SUBAPPLICATION INI_IN_AND_STORE_AUI2 (* INI Laden und Speichern von AUI2-Daten (reine Ganzzahl 0-N, kein Scale/Decimals) mit zusaetzlichem VALUEO (AUI, plain) fuer einen weiteren Consumer - analog INI_IN_AND_STORE_AUDI2, aber ueber den bidirektionalen AUI2-Adapter (UINT) statt AUDI2 (UDINT), z.B. fuer K eines AOption_AUI_DEMUX_N. *)
  (* Standard: 61499-2; Description: Copyright (c) 2026 Meisterschulen am Ostbahnhof This program and the accompanying materials are made available under the terms of the Eclipse Public License 2.0 which is available at https://www.eclipse.org/legal/epl-2.0/ SPDX-License-Identifier: EPL-2.0 *)
  (* Version 1.0, 2026-10-13, Franz Höpfinger, Meisterschulen am Ostbahnhof, UINT/AUI2-Pendant zu MyLib::sys::INI_IN_AND_STORE_AUDI2: NumericValue_IDA + AD_TO_AUI + AUI_TO_AUI2 + INI_AUI2 (bidirektionaler Adapter statt AUI+Split-Paar), AUI_TO_AUI2.AUI_OUT gesplittet auf Q_NumericValue_AUDI (VT-Anzeige, via AUI_TO_AUDI) und VALUEO (weiterer Consumer, z.B. AOption_AUI_DEMUX_N.K). Strukturell identisch zu INI_IN_AND_STORE_AUDI2, nur mit AUI2 statt AUDI2. *)
  PACKAGE MyLib::sys;
  IMPORT isobus::UT::Q::const::IDs::ID_NULL;
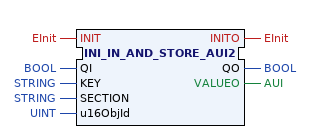
  EVENT_INPUT
    INIT : EInit; (* Initialization Request *)
  END_EVENT
  EVENT_OUTPUT
    INITO : EInit; (* Initialization Confirm *)
  END_EVENT
  VAR_INPUT
    QI : BOOL := TRUE; (* Quality Input - TRUE to enable service *)
    KEY : STRING; (* Key name. *)
    SECTION : STRING; (* Section name. *)
    u16ObjId : UINT := ID_NULL;
  END_VAR
  VAR_OUTPUT
    QO : BOOL; (* Quality Output - TRUE if service executed successfully *)
  END_VAR
  PLUGS
    VALUEO : adapter::types::unidirectional::AUI;
  END_PLUGS
  (* SETM=TRUE - der Boot-Wert laedt so oder so automatisch (INIT -> INITO -> GET -> GETO, unabhaengig von SETM). SETM=TRUE sorgt dafuer, dass auch eine LIVE-Aenderung waehrend des laufenden Betriebs sofort bestaetigt/zurueckgemeldet wird - wichtig, falls der frische Wert noch im selben Lauf weiterverwendet werden soll (z.B. hier ueber VALUEO). *)
  FBS
    ID : isobus::UT::io::NumericValue::NumericValue_IDA;
    AD_TO_AUI : adapter::conversion::unidirectional::AD_TO_AUI;
    AUI_TO_AUI2 : adapter::conversion::bidirectional::AUI_TO_AUI2;
    INI_AUI2 : eclipse4diac::storage::INI_AUI2(SETM := TRUE, DEFAULT_VALUE := UINT#0);
    AUI_SPLIT_2 : adapter::events::unidirectional::AUI_SPLIT_2;
    AUI_TO_AUDI : adapter::conversion::unidirectional::AUI_TO_AUDI;
    Q_NumericValue_AUDI : isobus::UT::Q::Q_NumericValue_AUDI;
    AND_QO : iec61131::booleanOperators::AND_BOOL_3;
  END_FBS
  EVENT_CONNECTIONS
    INIT TO ID.INIT;
    ID.INITO TO INI_AUI2.INIT;
    INI_AUI2.INITO TO Q_NumericValue_AUDI.INIT;
    Q_NumericValue_AUDI.INITO TO INITO;
    Q_NumericValue_AUDI.INITO TO AND_QO.REQ;
  END_CONNECTIONS
  DATA_CONNECTIONS
    KEY TO INI_AUI2.KEY;
    SECTION TO INI_AUI2.SECTION;
    u16ObjId TO ID.u16ObjId;
    u16ObjId TO Q_NumericValue_AUDI.u16ObjId;
    QI TO Q_NumericValue_AUDI.QI;
    QI TO ID.QI;
    QI TO INI_AUI2.QI;
    Q_NumericValue_AUDI.QO TO AND_QO.IN1;
    ID.QO TO AND_QO.IN2;
    INI_AUI2.QO TO AND_QO.IN3;
    AND_QO.OUT TO QO;
  END_CONNECTIONS
  ADAPTER_CONNECTIONS
    ID.IN TO AD_TO_AUI.AD_IN;
    AD_TO_AUI.AUI_OUT TO AUI_TO_AUI2.AUI_IN;
    AUI_TO_AUI2.AUI2_BIDIR TO INI_AUI2.VAL;
    AUI_TO_AUI2.AUI_OUT TO AUI_SPLIT_2.IN;
    AUI_SPLIT_2.OUT1 TO VALUEO;
    AUI_SPLIT_2.OUT2 TO AUI_TO_AUDI.AUI_IN;
    AUI_TO_AUDI.AUDI_OUT TO Q_NumericValue_AUDI.u32NewValue;
  END_CONNECTIONS
END_SUBAPPLICATION
